Fanuc KAREL source: KT00880.KL

PROGRAM KT00880
%NOLOCKGROUP
VAR
  I1: INTEGER
  I2: INTEGER
  OUT: INTEGER
BEGIN
  I1 = 2
  I2 = 3
  I1 = 2
  I2 = 3
  OUT = ATAN2(I1, I1)
END KT00880
